// Funzione M senza parametri: Nop, WaitH, LineNo, WaitStart.
FUNCTION F_MSimple : ST_MFuncDef
VAR_INPUT
	nChannel	: UINT;
	nMFunc		: UINT;
	eKind		: E_MFuncKind;
END_VAR

F_MSimple.nChannel := nChannel;
F_MSimple.nMFunc := nMFunc;
F_MSimple.eKind := eKind;

END_FUNCTION

(* stored: Version 1.1.0.1, ProductVersion 3.1.4024.12
   POU F_MSimple: Id {98606d1b-7ba3-46e8-9998-7505aa20ed5e}, SpecialFunc None *)
